Staubli VAL3: savePROG.pjx

--- savePROG.pjx ---
Parameters version=s8.10.3Cs9_BS2093 stackSize=5000 millimeterUnit=true
Data file=savePROG.dtx
Type name=progItem path=Disk://source/template/progItem/progItem.pjx

--- savePROG.dtx ---
public progItem pProgItem{}
  [Key1]
    progTemplate pProgTemplate
      [0]
        string sTRAJname
        num nType
        ifItem iIfItem
          [0]
            num nSigType[3]
            num nSigIndex[3]
            num nValue[3]
            bool bANDOR[2]
        switchItem sSwitchItem
          [0]
            num nSwitchValue
            string sIOValue
            bool bIOdisable
        forItem fForItem
          [0]
            num nLoopValue
            bool bIOdisable
            string sIOindex
